RoboDK station: Car_Painting_Cell_v2.rdk

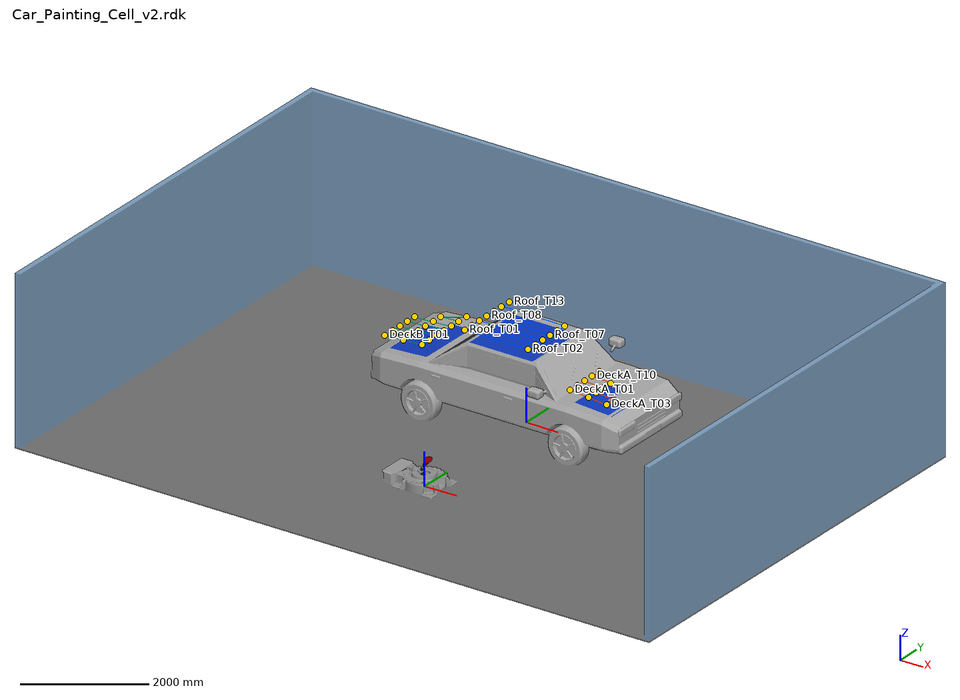
[picture v0: the station drawn from its stored meshes, robots at their saved joint values, targets as dots, program paths as lines]
Station Car_Painting_Cell_v2 (saved by RoboDK 6.1.1). Poses are relative to the parent item; angles as X-Y-Z fixed-axis rotations.
  - frame ABB IRB 6640-130/3.2 Base at (0, 0, 0) mm
    - robot ABB IRB 6640-130/3.2: 6 axes, payload 130 kg, reach 3200 mm, repeatability 0.05 mm, weight 1340 kg
        joint limits [-170, -65, -180, -300, -120, -360] to [170, 85, 70, 300, 120, 360]; home [0, 0, 0, 0, 0, 0]; saved at [119.913, 53.44, -52.284, 13.508, 41.833, -77.396]
      - tool Paint_Spray_Gun, TCP at (50, 0, 450) mm, rotated rx 0 ry 30 rz 0 deg, size 277.6 x 203.2 x 501.7 mm
  - Python program measure_car (listed below)
  - Python program build_cell (listed below)
  - object Floor at (0, 0, 0) mm, size 12000 x 8000 x 20 mm
  - object Wall_Back at (0, 0, 0) mm, size 12000 x 100 x 3000 mm
  - object Wall_Left at (0, 0, 0) mm, size 100 x 8000 x 3000 mm
  - object Wall_Right at (0, 0, 0) mm, size 100 x 8000 x 3000 mm
  - Python program reach_test (listed below)
  - Python program reach_test_roof (listed below)
  - frame Car_Frame at (0, 2750, 0) mm
    - object Car_Body at (0, 0, 0) mm, rotated rx 0 ry 0 rz 90 deg, size 2371.4 x 4800 x 1512.8 mm, geometry from Car_Body.stl
    - target Roof_T01 (Cartesian target) at (-566.92, -856.16, 1780.89) mm, rotated rx -140 ry 0 rz 0 deg; joints [69.061, 30.329, -32.85, 44.494, 71.837, -128.557] of ABB IRB 6640-130/3.2
    - target Roof_T02 (Cartesian target) at (629.09, -856.16, 1780.89) mm, rotated rx -140 ry 0 rz 0 deg; joints [69.061, 30.329, -32.85, 44.494, 71.837, -128.557] of ABB IRB 6640-130/3.2
    - target Roof_T03 (Cartesian target) at (629.09, -656.16, 1780.89) mm, rotated rx -140 ry 0 rz 0 deg; joints [69.061, 30.329, -32.85, 44.494, 71.837, -128.557] of ABB IRB 6640-130/3.2
    - target Roof_T04 (Cartesian target) at (-566.92, -656.16, 1780.89) mm, rotated rx -140 ry 0 rz 0 deg; joints [69.061, 30.329, -32.85, 44.494, 71.837, -128.557] of ABB IRB 6640-130/3.2
    - target Roof_T05 (Cartesian target) at (-566.92, -456.16, 1780.89) mm, rotated rx -140 ry 0 rz 0 deg; joints [69.061, 30.329, -32.85, 44.494, 71.837, -128.557] of ABB IRB 6640-130/3.2
    - target Roof_T06 (Cartesian target) at (629.09, -456.16, 1780.89) mm, rotated rx -140 ry 0 rz 0 deg; joints [69.061, 30.329, -32.85, 44.494, 71.837, -128.557] of ABB IRB 6640-130/3.2
    - target Roof_T07 (Cartesian target) at (629.09, -256.16, 1780.89) mm, rotated rx -140 ry 0 rz 0 deg; joints [69.061, 30.329, -32.85, 44.494, 71.837, -128.557] of ABB IRB 6640-130/3.2
    - target Roof_T08 (Cartesian target) at (-566.92, -256.16, 1780.89) mm, rotated rx -140 ry 0 rz 0 deg; joints [69.061, 30.329, -32.85, 44.494, 71.837, -128.557] of ABB IRB 6640-130/3.2
    - target Roof_T09 (Cartesian target) at (-566.92, -56.16, 1780.89) mm, rotated rx -140 ry 0 rz 0 deg; joints [69.061, 30.329, -32.85, 44.494, 71.837, -128.557] of ABB IRB 6640-130/3.2
    - target Roof_T10 (Cartesian target) at (629.09, -56.16, 1780.89) mm, rotated rx -140 ry 0 rz 0 deg; joints [69.061, 30.329, -32.85, 44.494, 71.837, -128.557] of ABB IRB 6640-130/3.2
    - target Roof_T11 (Cartesian target) at (629.09, 143.84, 1780.89) mm, rotated rx -140 ry 0 rz 0 deg; joints [69.061, 30.329, -32.85, 44.494, 71.837, -128.557] of ABB IRB 6640-130/3.2
    - target Roof_T12 (Cartesian target) at (-566.92, 143.84, 1780.89) mm, rotated rx -140 ry 0 rz 0 deg; joints [69.061, 30.329, -32.85, 44.494, 71.837, -128.557] of ABB IRB 6640-130/3.2
    - target Roof_T13 (Cartesian target) at (-566.92, 343.84, 1780.89) mm, rotated rx -140 ry 0 rz 0 deg; joints [69.061, 30.329, -32.85, 44.494, 71.837, -128.557] of ABB IRB 6640-130/3.2
    - target DeckA_T01 (Cartesian target) at (1400, -819.98, 1279.37) mm, rotated rx -140 ry 0 rz 0 deg; joints [0, 0, 0, 0, 0, 0] of ABB IRB 6640-130/3.2
    - target DeckA_T02 (Cartesian target) at (1750, -819.98, 1255.69) mm, rotated rx -140 ry 0 rz 0 deg; joints [0, 0, 0, 0, 0, 0] of ABB IRB 6640-130/3.2
    - target DeckA_T03 (Cartesian target) at (2100, -819.98, 1221.38) mm, rotated rx -140 ry 0 rz 0 deg; joints [0, 0, 0, 0, 0, 0] of ABB IRB 6640-130/3.2
    - target DeckA_T04 (Cartesian target) at (2100, -619.98, 1221.38) mm, rotated rx -140 ry 0 rz 0 deg; joints [0, 0, 0, 0, 0, 0] of ABB IRB 6640-130/3.2
    - target DeckA_T05 (Cartesian target) at (1750, -619.98, 1255.69) mm, rotated rx -140 ry 0 rz 0 deg; joints [0, 0, 0, 0, 0, 0] of ABB IRB 6640-130/3.2
    - target DeckA_T06 (Cartesian target) at (1400, -619.98, 1279.37) mm, rotated rx -140 ry 0 rz 0 deg; joints [0, 0, 0, 0, 0, 0] of ABB IRB 6640-130/3.2
    - target DeckA_T07 (Cartesian target) at (1400, -419.98, 1279.37) mm, rotated rx -140 ry 0 rz 0 deg; joints [0, 0, 0, 0, 0, 0] of ABB IRB 6640-130/3.2
    - target DeckA_T08 (Cartesian target) at (1750, -419.98, 1255.69) mm, rotated rx -140 ry 0 rz 0 deg; joints [0, 0, 0, 0, 0, 0] of ABB IRB 6640-130/3.2
    - target DeckA_T09 (Cartesian target) at (1750, -219.98, 1255.69) mm, rotated rx -140 ry 0 rz 0 deg; joints [0, 0, 0, 0, 0, 0] of ABB IRB 6640-130/3.2
    - target DeckA_T10 (Cartesian target) at (1400, -219.98, 1279.37) mm, rotated rx -140 ry 0 rz 0 deg; joints [0, 0, 0, 0, 0, 0] of ABB IRB 6640-130/3.2
    - target DeckA_T11 (Cartesian target) at (1400, -19.98, 1279.37) mm, rotated rx -140 ry 0 rz 0 deg; joints [0, 0, 0, 0, 0, 0] of ABB IRB 6640-130/3.2
    - target DeckB_T01 (Cartesian target) at (-2100, -819.98, 1240.33) mm, rotated rx -140 ry 0 rz 0 deg; joints [0, 0, 0, 0, 0, 0] of ABB IRB 6640-130/3.2
    - target DeckB_T02 (Cartesian target) at (-1750, -819.98, 1259.91) mm, rotated rx -140 ry 0 rz 0 deg; joints [0, 0, 0, 0, 0, 0] of ABB IRB 6640-130/3.2
    - target DeckB_T03 (Cartesian target) at (-1400, -819.98, 1279.49) mm, rotated rx -140 ry 0 rz 0 deg; joints [0, 0, 0, 0, 0, 0] of ABB IRB 6640-130/3.2
    - target DeckB_T04 (Cartesian target) at (-1400, -619.98, 1279.49) mm, rotated rx -140 ry 0 rz 0 deg; joints [0, 0, 0, 0, 0, 0] of ABB IRB 6640-130/3.2
    - target DeckB_T05 (Cartesian target) at (-1750, -619.98, 1259.91) mm, rotated rx -140 ry 0 rz 0 deg; joints [0, 0, 0, 0, 0, 0] of ABB IRB 6640-130/3.2
    - target DeckB_T06 (Cartesian target) at (-2100, -619.98, 1240.33) mm, rotated rx -140 ry 0 rz 0 deg; joints [0, 0, 0, 0, 0, 0] of ABB IRB 6640-130/3.2
    - target DeckB_T07 (Cartesian target) at (-2100, -419.98, 1240.33) mm, rotated rx -140 ry 0 rz 0 deg; joints [0, 0, 0, 0, 0, 0] of ABB IRB 6640-130/3.2
    - target DeckB_T08 (Cartesian target) at (-1750, -419.98, 1259.91) mm, rotated rx -140 ry 0 rz 0 deg; joints [0, 0, 0, 0, 0, 0] of ABB IRB 6640-130/3.2
    - target DeckB_T09 (Cartesian target) at (-1400, -419.98, 1279.49) mm, rotated rx -140 ry 0 rz 0 deg; joints [0, 0, 0, 0, 0, 0] of ABB IRB 6640-130/3.2
    - target DeckB_T10 (Cartesian target) at (-1400, -219.98, 1279.49) mm, rotated rx -140 ry 0 rz 0 deg; joints [0, 0, 0, 0, 0, 0] of ABB IRB 6640-130/3.2
    - target DeckB_T11 (Cartesian target) at (-1750, -219.98, 1259.91) mm, rotated rx -140 ry 0 rz 0 deg; joints [0, 0, 0, 0, 0, 0] of ABB IRB 6640-130/3.2
    - target DeckB_T12 (Cartesian target) at (-2100, -219.98, 1240.33) mm, rotated rx -140 ry 0 rz 0 deg; joints [0, 0, 0, 0, 0, 0] of ABB IRB 6640-130/3.2
    - target DeckB_T13 (Cartesian target) at (-2100, -19.98, 1240.33) mm, rotated rx -140 ry 0 rz 0 deg; joints [0, 0, 0, 0, 0, 0] of ABB IRB 6640-130/3.2
    - target DeckB_T14 (Cartesian target) at (-1750, -19.98, 1259.91) mm, rotated rx -140 ry 0 rz 0 deg; joints [0, 0, 0, 0, 0, 0] of ABB IRB 6640-130/3.2
    - target DeckB_T15 (Cartesian target) at (-1400, -19.98, 1279.49) mm, rotated rx -140 ry 0 rz 0 deg; joints [0, 0, 0, 0, 0, 0] of ABB IRB 6640-130/3.2
    - target DeckB_T16 (Cartesian target) at (-1400, 180.02, 1279.49) mm, rotated rx -140 ry 0 rz 0 deg; joints [0, 0, 0, 0, 0, 0] of ABB IRB 6640-130/3.2
    - target DeckB_T17 (Cartesian target) at (-1750, 180.02, 1259.91) mm, rotated rx -140 ry 0 rz 0 deg; joints [0, 0, 0, 0, 0, 0] of ABB IRB 6640-130/3.2
    - target DeckB_T18 (Cartesian target) at (-1400, 380.02, 1279.49) mm, rotated rx -140 ry 0 rz 0 deg; joints [0, 0, 0, 0, 0, 0] of ABB IRB 6640-130/3.2
  - Python program set_car_frame (listed below)
  - Python program make_roof_path (listed below)
  - program Paint_Roof (15 instructions, listed below)
  - Python program paint_roof_sim (listed below)
  - Python program make_deck_paths (listed below)
  - Python program check_mesh (listed below)
  - Python program check_heights (listed below)
  - program Paint_Deck_A (13 instructions, listed below)
  - program Paint_Deck_B (20 instructions, listed below)
  - Python program paint_all_sim (listed below)
  - object PaintStrip001 at (0, 0, 0) mm, size 299 x 200 x 0 mm
  - object PaintStrip002 at (0, 0, 0) mm, size 299 x 200 x 0 mm
  - object PaintStrip003 at (0, 0, 0) mm, size 299 x 200 x 0 mm
  - object PaintStrip004 at (0, 0, 0) mm, size 299 x 200 x 0 mm
  - object PaintStrip005 at (0, 0, 0) mm, size 299 x 200 x 0 mm
  - object PaintStrip006 at (0, 0, 0) mm, size 299 x 200 x 0 mm
  - object PaintStrip007 at (0, 0, 0) mm, size 299 x 200 x 0 mm
  - object PaintStrip008 at (0, 0, 0) mm, size 299 x 200 x 0 mm
  - object PaintStrip009 at (0, 0, 0) mm, size 299 x 200 x 0 mm
  - object PaintStrip010 at (0, 0, 0) mm, size 299 x 200 x 0 mm
  - object PaintStrip011 at (0, 0, 0) mm, size 299 x 200 x 0 mm
  - object PaintStrip012 at (0, 0, 0) mm, size 299 x 200 x 0 mm
  - object PaintStrip013 at (0, 0, 0) mm, size 299 x 200 x 0 mm
  - object PaintStrip014 at (0, 0, 0) mm, size 299 x 200 x 0 mm
  - object PaintStrip015 at (0, 0, 0) mm, size 299 x 200 x 0 mm
  - object PaintStrip016 at (0, 0, 0) mm, size 299 x 200 x 0 mm
  - object PaintStrip017 at (0, 0, 0) mm, size 299 x 200 x 0 mm
  - object PaintStrip018 at (0, 0, 0) mm, size 299 x 200 x 0 mm
  - object PaintStrip019 at (0, 0, 0) mm, size 299 x 200 x 0 mm
  - object PaintStrip020 at (0, 0, 0) mm, size 299 x 200 x 0 mm
  - object PaintStrip021 at (0, 0, 0) mm, size 299 x 200 x 0 mm
  - object PaintStrip022 at (0, 0, 0) mm, size 299 x 200 x 0 mm
  - object PaintStrip023 at (0, 0, 0) mm, size 299 x 200 x 0 mm
  - object PaintStrip024 at (0, 0, 0) mm, size 299 x 200 x 0 mm
  - object PaintStrip025 at (0, 0, 0) mm, size 87.5 x 200 x 5.9 mm
  - object PaintStrip026 at (0, 0, 0) mm, size 87.5 x 200 x 5.9 mm
  - object PaintStrip027 at (0, 0, 0) mm, size 87.5 x 200 x 5.9 mm
  - object PaintStrip028 at (0, 0, 0) mm, size 87.5 x 200 x 5.9 mm
  - object PaintStrip029 at (0, 0, 0) mm, size 87.5 x 200 x 5.9 mm
  - object PaintStrip030 at (0, 0, 0) mm, size 87.5 x 200 x 5.9 mm
  - object PaintStrip031 at (0, 0, 0) mm, size 87.5 x 200 x 5.9 mm
  - object PaintStrip032 at (0, 0, 0) mm, size 87.5 x 200 x 16.5 mm
  - object PaintStrip033 at (0, 0, 0) mm, size 87.5 x 200 x 16.5 mm
  - object PaintStrip034 at (0, 0, 0) mm, size 87.5 x 200 x 5.9 mm
  - object PaintStrip035 at (0, 0, 0) mm, size 87.5 x 200 x 5.9 mm
  - object PaintStrip036 at (0, 0, 0) mm, size 87.5 x 200 x 5.9 mm
  - object PaintStrip037 at (0, 0, 0) mm, size 87.5 x 200 x 5.9 mm
  - object PaintStrip038 at (0, 0, 0) mm, size 87.5 x 200 x 5.9 mm
  - object PaintStrip039 at (0, 0, 0) mm, size 87.5 x 200 x 5.9 mm
  - object PaintStrip040 at (0, 0, 0) mm, size 87.5 x 200 x 5.9 mm
  - object PaintStrip041 at (0, 0, 0) mm, size 87.5 x 200 x 5.9 mm
  - object PaintStrip042 at (0, 0, 0) mm, size 87.5 x 200 x 5.9 mm
  - object PaintStrip043 at (0, 0, 0) mm, size 87.5 x 200 x 5.9 mm
  - object PaintStrip044 at (0, 0, 0) mm, size 87.5 x 200 x 5.9 mm
  - object PaintStrip045 at (0, 0, 0) mm, size 87.5 x 200 x 5.9 mm
  - object PaintStrip046 at (0, 0, 0) mm, size 87.5 x 200 x 5.9 mm
  - object PaintStrip047 at (0, 0, 0) mm, size 87.5 x 200 x 5.9 mm
  - object PaintStrip048 at (0, 0, 0) mm, size 87.5 x 200 x 5.9 mm
  - object PaintStrip049 at (0, 0, 0) mm, size 87.5 x 200 x 4.9 mm
  - object PaintStrip050 at (0, 0, 0) mm, size 87.5 x 200 x 4.9 mm
  - object PaintStrip051 at (0, 0, 0) mm, size 87.5 x 200 x 4.9 mm
  - object PaintStrip052 at (0, 0, 0) mm, size 87.5 x 200 x 4.9 mm
  - object PaintStrip053 at (0, 0, 0) mm, size 87.5 x 200 x 4.9 mm
  - object PaintStrip054 at (0, 0, 0) mm, size 87.5 x 200 x 4.9 mm
  - object PaintStrip055 at (0, 0, 0) mm, size 87.5 x 200 x 4.9 mm
  - object PaintStrip056 at (0, 0, 0) mm, size 87.5 x 200 x 4.9 mm
  - object PaintStrip057 at (0, 0, 0) mm, size 87.5 x 200 x 4.9 mm
  - object PaintStrip058 at (0, 0, 0) mm, size 87.5 x 200 x 4.9 mm
  - object PaintStrip059 at (0, 0, 0) mm, size 87.5 x 200 x 4.9 mm
  - object PaintStrip060 at (0, 0, 0) mm, size 87.5 x 200 x 4.9 mm
  - object PaintStrip061 at (0, 0, 0) mm, size 87.5 x 200 x 4.9 mm
  - object PaintStrip062 at (0, 0, 0) mm, size 87.5 x 200 x 4.9 mm
  - object PaintStrip063 at (0, 0, 0) mm, size 87.5 x 200 x 4.9 mm
  - object PaintStrip064 at (0, 0, 0) mm, size 87.5 x 200 x 4.9 mm
  - object PaintStrip065 at (0, 0, 0) mm, size 87.5 x 200 x 4.9 mm
  - object PaintStrip066 at (0, 0, 0) mm, size 87.5 x 200 x 4.9 mm
  - object PaintStrip067 at (0, 0, 0) mm, size 87.5 x 200 x 4.9 mm
  - object PaintStrip068 at (0, 0, 0) mm, size 87.5 x 200 x 4.9 mm
  - object PaintStrip069 at (0, 0, 0) mm, size 87.5 x 200 x 4.9 mm
  - object PaintStrip070 at (0, 0, 0) mm, size 87.5 x 200 x 4.9 mm
  - object PaintStrip071 at (0, 0, 0) mm, size 87.5 x 200 x 4.9 mm
  - object PaintStrip072 at (0, 0, 0) mm, size 87.5 x 200 x 4.9 mm
  - object PaintStrip073 at (0, 0, 0) mm, size 87.5 x 200 x 4.9 mm
  - object PaintStrip074 at (0, 0, 0) mm, size 87.5 x 200 x 4.9 mm
  - object PaintStrip075 at (0, 0, 0) mm, size 87.5 x 200 x 4.9 mm
  - object PaintStrip076 at (0, 0, 0) mm, size 87.5 x 200 x 4.9 mm
  - object PaintStrip077 at (0, 0, 0) mm, size 87.5 x 200 x 4.9 mm
  - object PaintStrip078 at (0, 0, 0) mm, size 87.5 x 200 x 4.9 mm
  - object PaintStrip079 at (0, 0, 0) mm, size 87.5 x 200 x 4.9 mm
  - object PaintStrip080 at (0, 0, 0) mm, size 87.5 x 200 x 4.9 mm
  - object PaintStrip081 at (0, 0, 0) mm, size 87.5 x 200 x 4.9 mm
  - object PaintStrip082 at (0, 0, 0) mm, size 87.5 x 200 x 4.9 mm
  - object PaintStrip083 at (0, 0, 0) mm, size 87.5 x 200 x 4.9 mm
  - object PaintStrip084 at (0, 0, 0) mm, size 87.5 x 200 x 4.9 mm
  - object PaintStrip085 at (0, 0, 0) mm, size 87.5 x 200 x 4.9 mm
  - object PaintStrip086 at (0, 0, 0) mm, size 87.5 x 200 x 4.9 mm
  - object PaintStrip087 at (0, 0, 0) mm, size 87.5 x 200 x 4.9 mm
  - object PaintStrip088 at (0, 0, 0) mm, size 87.5 x 200 x 4.9 mm
  - object PaintStrip089 at (0, 0, 0) mm, size 87.5 x 200 x 4.9 mm
  - object PaintStrip090 at (0, 0, 0) mm, size 87.5 x 200 x 4.9 mm
  - object PaintStrip091 at (0, 0, 0) mm, size 87.5 x 200 x 4.9 mm
  - object PaintStrip092 at (0, 0, 0) mm, size 87.5 x 200 x 4.9 mm
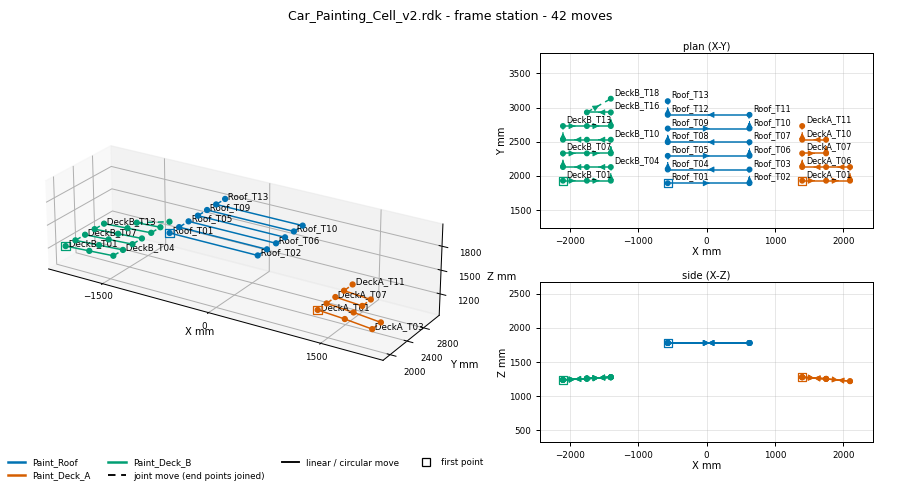
[picture p0: tool path of Car_Painting_Cell_v2.rdk in frame station, 42 of 42 moves have a stored position in this frame; points joined in program order, loops and branches not executed]

--- Python program measure_car ---
from robodk.robolink import *
from robodk.robomath import *
import numpy as np

RDK = Robolink()
car = RDK.Item('Car_Body')

# 1) scale uniformly so the long side (local Y) is 4800 mm
pts, _ = car.GetPoints(FEATURE_OBJECT_MESH)
p = np.array(pts)[:, :3]
length = p[:, 1].max() - p[:, 1].min()
car.Scale(4800.0 / length)

# 2) re-read the scaled mesh and rotate 90 deg about Z (x,y) -> (-y,x)
pts, _ = car.GetPoints(FEATURE_OBJECT_MESH)
p = np.array(pts)[:, :3]
rx, ry, rz = -p[:, 1], p[:, 0], p[:, 2]

# 3) centre the car in X, put its centreline 2300 mm from the robot base, wheels on Z=0
tx = -(rx.min() + rx.max()) / 2
ty = 2300 - (ry.min() + ry.max()) / 2
tz = -rz.min()
car.setPose(transl(tx, ty, tz) * rotz(pi / 2))

# 4) light grey colour (R,G,B,A from 0 to 1)
car.setColor([0.8, 0.8, 0.8, 1.0])

RDK.ShowMessage("Car size X,Y,Z = %.0f x %.0f x %.0f mm\nPlaced at X=%.0f Y=%.0f Z=%.0f" %
                (rx.max() - rx.min(), ry.max() - ry.min(), rz.max() - rz.min(), tx, ty, tz), True)

--- Python program build_cell ---
from robodk.robolink import *

RDK = Robolink()

def box(x0, x1, y0, y1, z0, z1):
    """12 triangles of an axis-aligned box, as a flat list of vertices."""
    v = [[x0,y0,z0],[x1,y0,z0],[x1,y1,z0],[x0,y1,z0],
         [x0,y0,z1],[x1,y0,z1],[x1,y1,z1],[x0,y1,z1]]
    faces = [(0,2,1),(0,3,2),(4,5,6),(4,6,7),(0,1,5),(0,5,4),
             (1,2,6),(1,6,5),(2,3,7),(2,7,6),(3,0,4),(3,4,7)]
    return [v[i] for f in faces for i in f]

# remove old objects if the script is run again
for name in ['Floor', 'Wall_Back', 'Wall_Left', 'Wall_Right']:
    old = RDK.Item(name)
    if old.Valid():
        old.Delete()

# 12 m x 8 m floor, top surface at Z = 0, robot base at (0,0,0)
floor = RDK.AddShape(box(-6000, 6000, -2500, 5500, -20, 0))
floor.setName('Floor')
floor.setColor([0.55, 0.55, 0.55, 1.0])

# 3 m high translucent walls: back and both ends (front left open for the camera)
wall_color = [0.6, 0.75, 0.9, 0.3]
w1 = RDK.AddShape(box(-6000, 6000, 5400, 5500, 0, 3000))
w1.setName('Wall_Back');  w1.setColor(wall_color)
w2 = RDK.AddShape(box(-6000, -5900, -2500, 5500, 0, 3000))
w2.setName('Wall_Left');  w2.setColor(wall_color)
w3 = RDK.AddShape(box(5900, 6000, -2500, 5500, 0, 3000))
w3.setName('Wall_Right'); w3.setColor(wall_color)

RDK.ShowMessage('Cell built: floor 12000 x 8000 mm, walls 3000 mm high', True)

--- Python program reach_test ---
from robodk.robolink import *
from robodk.robomath import *
import numpy as np

RDK = Robolink()
robot = RDK.Item('ABB IRB 6640-130/3.2')
car = RDK.Item('Car_Body')
tool = RDK.Item('Paint_Spray_Gun')

# car bounding box in station coordinates
pts, _ = car.GetPoints(FEATURE_OBJECT_MESH)
p = np.array(pts)[:, :3]
T = np.array(car.Pose().rows)
w = (T[:3, :3] @ p.T).T + T[:3, 3]
mn, mx = w.min(axis=0), w.max(axis=0)
cy = (mn[1] + mx[1]) / 2
stand = 250  # gun distance from the surface, mm

def mk(pos, x, y, z):
    return Mat([[x[0], y[0], z[0], pos[0]],
                [x[1], y[1], z[1], pos[1]],
                [x[2], y[2], z[2], pos[2]],
                [0, 0, 0, 1]])

def reachable(pose):
    try:
        j = robot.SolveIK(pose, tool=tool.PoseTool())
        return len(j.list()) == 6
    except Exception:
        return False

xs = list(range(-2400, 2401, 400))
zs = 0.6 * mx[2]
tests = {
    'Top (gun pointing down)': [mk([x, cy, mx[2] + stand], [1,0,0], [0,-1,0], [0,0,-1]) for x in xs],
    'Near side (gun pointing +Y)': [mk([x, mn[1] - stand, zs], [1,0,0], [0,0,-1], [0,1,0]) for x in xs],
    'Far side (gun pointing -Y)': [mk([x, mx[1] + stand, zs], [1,0,0], [0,0,1], [0,-1,0]) for x in xs],
}

msg = "Car size: %.0f x %.0f x %.0f mm\n" % tuple(mx - mn)
for name, poses in tests.items():
    ok = [reachable(P) for P in poses]
    bad = [xs[i] for i, o in enumerate(ok) if not o]
    msg += "\n%s: %d of %d reachable" % (name, sum(ok), len(ok))
    if bad:
        msg += "\n   NOT reachable at X = %s" % bad
RDK.ShowMessage(msg, True)

--- Python program reach_test_roof ---
from robodk.robolink import *
from robodk.robomath import *
import numpy as np

RDK = Robolink()
robot = RDK.Item('ABB IRB 6640-130/3.2')
car = RDK.Item('Car_Body')
tool = RDK.Item('Paint_Spray_Gun')

pts, _ = car.GetPoints(FEATURE_OBJECT_MESH)
p = np.array(pts)[:, :3]
T = np.array(car.PoseAbs().rows)
w = (T[:3, :3] @ p.T).T + T[:3, 3]
mn, mx = w.min(axis=0), w.max(axis=0)
cy = (mn[1] + mx[1]) / 2
top = mx[2]
stand = 250  # mm

def pose_for(P, tilt_deg):
    t = np.radians(tilt_deg)
    s, c = np.sin(t), np.cos(t)
    d = np.array([0, s, -c])      # spray direction: down, leaning away from the robot (+Y)
    x = np.array([1, 0, 0])
    y = np.cross(d, x)
    pos = np.array(P) - stand * d
    return Mat([[x[0], y[0], d[0], pos[0]],
                [x[1], y[1], d[1], pos[1]],
                [x[2], y[2], d[2], pos[2]],
                [0, 0, 0, 1]])

def reachable(pose):
    try:
        j = robot.SolveIK(pose, tool=tool.PoseTool())
        return len(j.list()) == 6
    except Exception:
        return False

xs = list(range(-2000, 2001, 400))
msg = "Roof-height points, car Y = %.0f mm (13... %d points per row)\n" % (cy, len(xs))
for tilt in [0, 20, 40]:
    msg += "\nTilt %d deg:" % tilt
    for dy in [-600, -300, 0]:
        n = sum(reachable(pose_for([x, cy + dy, top], tilt)) for x in xs)
        msg += "\n   %4d mm from centreline: %d of %d" % (dy, n, len(xs))
RDK.ShowMessage(msg, True)

--- Python program set_car_frame ---
from robodk.robolink import *
from robodk.robomath import *

RDK = Robolink()
frame = RDK.Item('Car_Frame')
frame.setPose(transl(0, 2750, 0))
p = frame.Pose().Pos()
RDK.ShowMessage("Car_Frame is now at X=%.0f Y=%.0f Z=%.0f" % (p[0], p[1], p[2]), True)

--- Python program make_roof_path ---
from robodk.robolink import *
from robodk.robomath import *
import numpy as np

RDK = Robolink()
robot = RDK.Item('ABB IRB 6640-130/3.2')
car = RDK.Item('Car_Body')
tool = RDK.Item('Paint_Spray_Gun')
frame = RDK.Item('Car_Frame')

# delete old roof targets/program if the script is run again
for it in RDK.ItemList(ITEM_TYPE_TARGET):
    if it.Name().startswith('Roof_'):
        it.Delete()
old = RDK.Item('Paint_Roof')
if old.Valid():
    old.Delete()

# car mesh in station coordinates
pts, _ = car.GetPoints(FEATURE_OBJECT_MESH)
p = np.array(pts)[:, :3]
T = np.array(car.PoseAbs().rows)
w = (T[:3, :3] @ p.T).T + T[:3, 3]
top = w[:, 2].max()

# flat roof area = points within 60 mm of the highest point
roof = w[w[:, 2] > top - 60]
x0, x1 = roof[:, 0].min() + 50, roof[:, 0].max() - 50
y0, y1 = roof[:, 1].min() + 50, roof[:, 1].max() - 50

stand = 350      # gun distance from the surface, mm
tilt = 40        # degrees, leaning away from the robot
spacing = 200    # distance between stripes, mm
t = np.radians(tilt)
d = np.array([0, np.sin(t), -np.cos(t)])   # spray direction
xa = np.array([1.0, 0, 0])
ya = np.cross(d, xa)

def abs_pose(x, y):
    pos = np.array([x, y, top]) - stand * d
    return Mat([[xa[0], ya[0], d[0], pos[0]],
                [xa[1], ya[1], d[1], pos[1]],
                [xa[2], ya[2], d[2], pos[2]],
                [0, 0, 0, 1]])

def reachable(P):
    try:
        return len(robot.SolveIK(P, tool=tool.PoseTool()).list()) == 6
    except Exception:
        return False

prog = RDK.AddProgram('Paint_Roof', robot)
prog.setPoseFrame(frame)
prog.setPoseTool(tool)
inv_frame = frame.PoseAbs().inv()

ys = np.arange(y0, y1 + 1, spacing)
n_ok, n_bad, k = 0, 0, 0
for i, y in enumerate(ys):
    xs = [x0, x1] if i % 2 == 0 else [x1, x0]   # zig-zag
    for j, x in enumerate(xs):
        P = abs_pose(x, y)
        if not reachable(P):
            n_bad += 1
            continue
        k += 1
        tg = RDK.AddTarget('Roof_T%02d' % k, frame, robot)
        tg.setAsCartesianTarget()
        tg.setPose(inv_frame * P)
        if n_ok == 0 or j == 0:
            prog.MoveJ(tg)
        else:
            prog.MoveL(tg)
        n_ok += 1

RDK.ShowMessage("Roof: %.0f x %.0f mm, %d stripes\nTargets created: %d, unreachable (skipped): %d"
                % (x1 - x0, y1 - y0, len(ys), n_ok, n_bad), True)

--- program Paint_Roof (robot ABB IRB 6640-130/3.2) ---
  Set Ref.: Car_Frame
  Set Tool: Paint_Spray_Gun
  MoveJ (Roof_T01)
  MoveL (Roof_T02)
  MoveJ (Roof_T03)
  MoveL (Roof_T04)
  MoveJ (Roof_T05)
  MoveL (Roof_T06)
  MoveJ (Roof_T07)
  MoveL (Roof_T08)
  MoveJ (Roof_T09)
  MoveL (Roof_T10)
  MoveJ (Roof_T11)
  MoveL (Roof_T12)
  MoveJ (Roof_T13)

--- Python program paint_roof_sim ---
from robodk.robolink import *

RDK = Robolink()
robot = RDK.Item('ABB IRB 6640-130/3.2')
tool = RDK.Item('Paint_Spray_Gun')
car = RDK.Item('Car_Body')
frame = RDK.Item('Car_Frame')
robot.setPoseFrame(frame)
robot.setPoseTool(tool)

RDK.Spray_Clear()
RDK.Spray_Add(tool, car)
RDK.Spray_SetState(SPRAY_OFF)

targets = sorted([t for t in RDK.ItemList(ITEM_TYPE_TARGET) if t.Name().startswith('DeckB_T')],
                 key=lambda t: t.Name())
robot.MoveJ(targets[0])
RDK.Spray_SetState(SPRAY_ON)
for t in targets[1:4]:
    robot.MoveL(t)
RDK.Spray_SetState(SPRAY_OFF)
RDK.ShowMessage('Test done', True)

--- Python program make_deck_paths ---
from robodk.robolink import *
from robodk.robomath import *
import numpy as np

RDK = Robolink()
robot = RDK.Item('ABB IRB 6640-130/3.2')
tool = RDK.Item('Paint_Spray_Gun')
frame = RDK.Item('Car_Frame')

# park the arm away from the car so the height probe hits only the car
robot.setJoints([0, 0, 0, 0, 0, 0])

# delete old deck targets and programs
for it in RDK.ItemList(ITEM_TYPE_TARGET):
    if it.Name().startswith('DeckA_') or it.Name().startswith('DeckB_'):
        it.Delete()
for n in ['Paint_Deck_A', 'Paint_Deck_B']:
    old = RDK.Item(n)
    if old.Valid():
        old.Delete()

cy = 2755
stand, tilt = 350, 40
t = np.radians(tilt)
d = np.array([0, np.sin(t), -np.cos(t)])
xa = np.array([1.0, 0, 0])
ya = np.cross(d, xa)

def surf(x, y):
    hit, item, xyz = RDK.Collision_Line([x, y, 3000], [x, y, 0])
    if hit and item.Name() == 'Car_Body':
        return xyz[2]
    return None

def abs_pose(x, y, z):
    pos = np.array([x, y, z]) - stand * d
    return Mat([[xa[0], ya[0], d[0], pos[0]],
                [xa[1], ya[1], d[1], pos[1]],
                [xa[2], ya[2], d[2], pos[2]],
                [0, 0, 0, 1]])

def reachable(P):
    try:
        return len(robot.SolveIK(P, tool=tool.PoseTool()).list()) == 6
    except Exception:
        return False

inv_frame = frame.PoseAbs().inv()
zones = [('A', 1400, 2100), ('B', -2100, -1400)]
ys = np.linspace(cy - 600, cy + 600, 7)
msg = ''
for tag, xlo, xhi in zones:
    prog = RDK.AddProgram('Paint_Deck_' + tag, robot)
    prog.setPoseFrame(frame)
    prog.setPoseTool(tool)
    k, bad, zmin, zmax = 0, 0, 9999, 0
    for i, y in enumerate(ys):
        xs = [xlo, (xlo + xhi) / 2, xhi]
        if i % 2 == 1:
            xs = xs[::-1]
        first = True
        for x in xs:
            z = surf(x, y)
            if z is None:
                bad += 1
                continue
            P = abs_pose(x, y, z)
            if not reachable(P):
                bad += 1
                continue
            k += 1
            zmin, zmax = min(zmin, z), max(zmax, z)
            tg = RDK.AddTarget('Deck%s_T%02d' % (tag, k), frame, robot)
            tg.setAsCartesianTarget()
            tg.setPose(inv_frame * P)
            tg.setVisible(False)
            if first:
                prog.MoveJ(tg)
                first = False
            else:
                prog.MoveL(tg)
    msg += "End %s: X %d to %d\n   surface Z %.0f to %.0f\n   targets %d, skipped %d\n" % (
        tag, xlo, xhi, zmin, zmax, k, bad)

RDK.ShowMessage(msg, True)

--- Python program check_mesh ---
from robodk.robolink import *
import numpy as np

RDK = Robolink()
car = RDK.Item('Car_Body')
pts, _ = car.GetPoints(FEATURE_OBJECT_MESH)
a = np.array(pts)
T = np.array(car.PoseAbs().rows)
w = (T[:3, :3] @ a[:, :3].T).T + T[:3, 3]

cy = (w[:, 1].min() + w[:, 1].max()) / 2

def zr(x0, x1):
    inx = (w[:, 0] > x0) & (w[:, 0] < x1)
    near = abs(w[:, 1] - cy) < 700
    s = w[inx & near]
    if len(s) == 0:
        return "no points"
    return "%d pts, Z %.0f to %.0f" % (len(s), s[:, 2].min(), s[:, 2].max())

msg = "Total points: %d\n" % len(a)
for x0 in range(-2400, 2400, 400):
    msg += "X %5d..%5d: %s\n" % (x0, x0 + 400, zr(x0, x0 + 400))
RDK.ShowMessage(msg, True)

--- Python program check_heights ---
from robodk.robolink import *
from robodk.robomath import *
import numpy as np

RDK = Robolink()
RDK.setCollisionActive(COLLISION_ON)
robot = RDK.Item('ABB IRB 6640-130/3.2')
tool = RDK.Item('Paint_Spray_Gun')
home = [0, 0, 0, 0, 0, 0]
robot.setJoints(home)   # park arm so the height probe only hits the car

cy, stand = 2755, 350

def surf(x, y):
    hit, item, xyz = RDK.Collision_Line([x, y, 3000], [x, y, 0])
    if hit and item.Name() == 'Car_Body':
        return xyz[2]
    return None

def pose(x, y, z, a, b):
    a, b = np.radians(a), np.radians(b)
    d = np.array([np.sin(a), np.sin(b)*np.cos(a), -np.cos(a)*np.cos(b)])
    ya = np.cross(d, [1.0, 0, 0]); ya /= np.linalg.norm(ya)
    xa = np.cross(ya, d)
    p = np.array([x, y, z]) - stand * d
    return Mat([[xa[0], ya[0], d[0], p[0]],
                [xa[1], ya[1], d[1], p[1]],
                [xa[2], ya[2], d[2], p[2]],
                [0, 0, 0, 1]])

def status(P):
    # returns 0 = unreachable, 1 = reachable but every solution collides, 2 = reachable and collision-free
    try:
        sols = robot.SolveIK_All(P, tool.PoseTool())
        cols = sols.Cols()
    except Exception:
        return 0
    cols = [c for c in cols if len(c) >= 6]
    if not cols:
        return 0
    for c in cols:
        robot.setJoints(c[:6])
        if RDK.Collisions() == 0:
            return 2
    return 1

zones = [('A', 1400, 2100), ('B', -2100, -1400)]
ys = np.linspace(cy - 600, cy + 600, 7)
tilts = [(0, 40), (0, -40), (0, 0), (40, 0), (-40, 0), (30, 30), (-30, 30)]
msg = ''
for tag, xlo, xhi in zones:
    msg += 'End %s (of 21 points)\n' % tag
    for (a, b) in tilts:
        c = [0, 0, 0]
        for y in ys:
            for x in [xlo, (xlo + xhi) / 2, xhi]:
                z = surf(x, y)
                if z is None:
                    continue
                c[status(pose(x, y, z, a, b))] += 1
        msg += '  tilt(%d,%d): OK %d | collide %d | unreachable %d\n' % (a, b, c[2], c[1], c[0])
robot.setJoints(home)
RDK.ShowMessage(msg, True)

--- program Paint_Deck_A (robot ABB IRB 6640-130/3.2) ---
  Set Ref.: Car_Frame
  Set Tool: Paint_Spray_Gun
  MoveJ (DeckA_T01)
  MoveL (DeckA_T02)
  MoveL (DeckA_T03)
  MoveJ (DeckA_T04)
  MoveL (DeckA_T05)
  MoveL (DeckA_T06)
  MoveJ (DeckA_T07)
  MoveL (DeckA_T08)
  MoveJ (DeckA_T09)
  MoveL (DeckA_T10)
  MoveJ (DeckA_T11)

--- program Paint_Deck_B (robot ABB IRB 6640-130/3.2) ---
  Set Ref.: Car_Frame
  Set Tool: Paint_Spray_Gun
  MoveJ (DeckB_T01)
  MoveL (DeckB_T02)
  MoveL (DeckB_T03)
  MoveJ (DeckB_T04)
  MoveL (DeckB_T05)
  MoveL (DeckB_T06)
  MoveJ (DeckB_T07)
  MoveL (DeckB_T08)
  MoveL (DeckB_T09)
  MoveJ (DeckB_T10)
  MoveL (DeckB_T11)
  MoveL (DeckB_T12)
  MoveJ (DeckB_T13)
  MoveL (DeckB_T14)
  MoveL (DeckB_T15)
  MoveJ (DeckB_T16)
  MoveL (DeckB_T17)
  MoveJ (DeckB_T18)

--- Python program paint_all_sim ---
from robodk.robolink import *
from robodk.robomath import *
import numpy as np

RDK = Robolink()
robot = RDK.Item('ABB IRB 6640-130/3.2')
tool = RDK.Item('Paint_Spray_Gun')
car = RDK.Item('Car_Body')
frame = RDK.Item('Car_Frame')

frame.setPose(transl(0, 2750, 0))

for it in RDK.ItemList(ITEM_TYPE_OBJECT):
    if it.Name().startswith('PaintStrip'):
        it.Delete()

robot.setJoints([0, 0, 0, 0, 0, 0])   # park the arm so the height probe hits only the car

def surf(x, y):
    hit, item, xyz = RDK.Collision_Line([x, y, 3000], [x, y, 0])
    if hit and item.Name() == 'Car_Body':
        return xyz[2]
    return None

def seg_tris(x0, x1, y, half=100):
    za, zb = surf(x0, y), surf(x1, y)
    if za is None or zb is None:
        return []
    a = [x0, y - half, za + 3]
    b = [x1, y - half, zb + 3]
    c = [x1, y + half, zb + 3]
    d = [x0, y + half, za + 3]
    return [a, b, c, a, c, d]

N = 4                                   # pieces of paint per stripe segment
dy = 350 * np.sin(np.radians(40))

# step 1: build the plan (poses along each stripe + the paint piece under each)
plan = []
for prefix in ['Roof_T', 'DeckA_T', 'DeckB_T']:
    targets = sorted([t for t in RDK.ItemList(ITEM_TYPE_TARGET) if t.Name().startswith(prefix)],
                     key=lambda t: t.Name())
    ys = [t.Pose().Pos()[1] for t in targets]
    i = 0
    while i < len(targets):
        j = i + 1
        while j < len(targets) and abs(ys[j] - ys[i]) < 1:
            j += 1
        if j - i >= 2:
            steps = []
            for k in range(i, j - 1):
                ta, tb = targets[k], targets[k + 1]
                Pa, Pb = ta.Pose(), tb.Pose()
                va = np.array(Pa.Pos())
                vb = np.array(Pb.Pos())
                aa = np.array(ta.PoseAbs().Pos())
                ab = np.array(tb.PoseAbs().Pos())
                for s in range(N):
                    f0, f1 = s / N, (s + 1) / N
                    d1 = (vb - va) * f1
                    pose = transl(d1[0], d1[1], d1[2]) * Pa
                    x0 = aa[0] + (ab[0] - aa[0]) * f0
                    x1 = aa[0] + (ab[0] - aa[0]) * f1
                    steps.append((pose, seg_tris(x0, x1, aa[1] + dy)))
            plan.append((targets[i], steps))
        i = j

# step 2: paint
robot.setPoseFrame(frame)
robot.setPoseTool(tool)
RDK.Spray_Clear()
RDK.Spray_Add(tool, car)
RDK.Spray_SetState(SPRAY_OFF)

n, skipped = 0, 0
for start, steps in plan:
    try:
        robot.MoveJ(start)
    except Exception:
        skipped += 1
        continue
    RDK.Spray_SetState(SPRAY_ON)
    for pose, tris in steps:
        try:
            robot.MoveL(pose)
        except Exception:
            break
        if tris:
            n += 1
            s = RDK.AddShape(tris)
            s.setName('PaintStrip%03d' % n)
            s.setColor([0.1, 0.3, 0.9, 1.0])   # blue paint
    RDK.Spray_SetState(SPRAY_OFF)

RDK.ShowMessage('Painting finished. Blue paint pieces: %d, stripes skipped: %d' % (n, skipped), True)
